FUNCTION_BLOCK SKILL_RunLogic (* The state machine of SKILL_Run: the precondition, waiting for the equipment, the command, the end condition, the timeout, the closing command. Technical: One run of a skill primitive: Pre, then the equipment free (0.5 s grace), Command until Post or the timer (Timed), Inv over it, StopCommand at the end, played before the end is reported *)
  (* Standard: 61499-2 *)
  (* Version 0.1, 2026-09-28, Project contributors, AAU Smart Production Lab *)
  PACKAGE modlib;
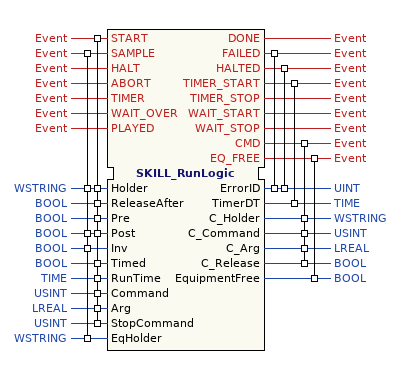
  EVENT_INPUT
    START WITH Holder, ReleaseAfter, Pre, Post, Timed, RunTime, Command, Arg, StopCommand; (* Start the run with what the contract says (Pre first) *)
    SAMPLE WITH Holder, Post, Inv, EqHolder; (* The equipment's newest state, as the contract judges it (Post, Inv, EqHolder) *)
    HALT; (* Stop the run (ErrorID Interrupted) *)
    ABORT; (* Abort the run: the equipment off and given up *)
    TIMER; (* The run's timer expired *)
    WAIT_OVER; (* Waited long enough for another holder to let go *)
    PLAYED; (* The command's phases were played *)
  END_EVENT
  EVENT_OUTPUT
    DONE; (* The run succeeded *)
    FAILED WITH ErrorID; (* The run failed (ErrorID) *)
    HALTED WITH ErrorID; (* The run was stopped *)
    TIMER_START WITH TimerDT; (* Start the timer (TimerDT) *)
    TIMER_STOP; (* Stop the timer *)
    WAIT_START; (* Start waiting for the equipment *)
    WAIT_STOP; (* Stop waiting *)
    CMD WITH C_Holder, C_Command, C_Arg, C_Release; (* Send a command to the equipment *)
    EQ_FREE WITH EquipmentFree; (* EquipmentFree is updated *)
  END_EVENT
  VAR_INPUT
    Holder : WSTRING; (* The name the equipment is held under: the skill's own, or for a step the skill it belongs to *)
    ReleaseAfter : BOOL; (* Give up the equipment with the run's last command *)
    Pre : BOOL; (* The precondition holds: the run may start (else PreconditionViolated, 1) *)
    Post : BOOL; (* The postcondition holds: the skill is done *)
    Inv : BOOL := TRUE; (* The invariant holds: the run may go on (else InvariantViolated, 2) *)
    Timed : BOOL; (* The skill ends after RunTime (TRUE), or when Post holds, failing after RunTime (FALSE) *)
    RunTime : TIME; (* How long it runs (Timed), or may take before it fails with Timeout (3) *)
    Command : USINT; (* The command's code to send while it runs *)
    Arg : LREAL; (* The command's argument (e.g. a position) *)
    StopCommand : USINT; (* The command's code to send when it is done or halted *)
    EqHolder : WSTRING; (* Who holds the equipment now (empty: free) *)
  END_VAR
  VAR_OUTPUT
    ErrorID : UINT; (* Error code: 0 none, 1 PreconditionViolated, 2 InvariantViolated, 3 Timeout, 4 NotReady, 5 NotPermitted, 6 Busy, 7 Interrupted, 8 OutOfRange *)
    TimerDT : TIME; (* How long the timer runs *)
    C_Holder : WSTRING; (* Sent with the command: who holds the equipment *)
    C_Command : USINT; (* Sent with the command: the command's code *)
    C_Arg : LREAL; (* Sent with the command: its argument (e.g. a position) *)
    C_Release : BOOL; (* Sent with the command: give up the equipment after it *)
    EquipmentFree : BOOL; (* The equipment is free, or held under Holder *)
  END_VAR
  VAR
    Outcome : USINT;
  END_VAR
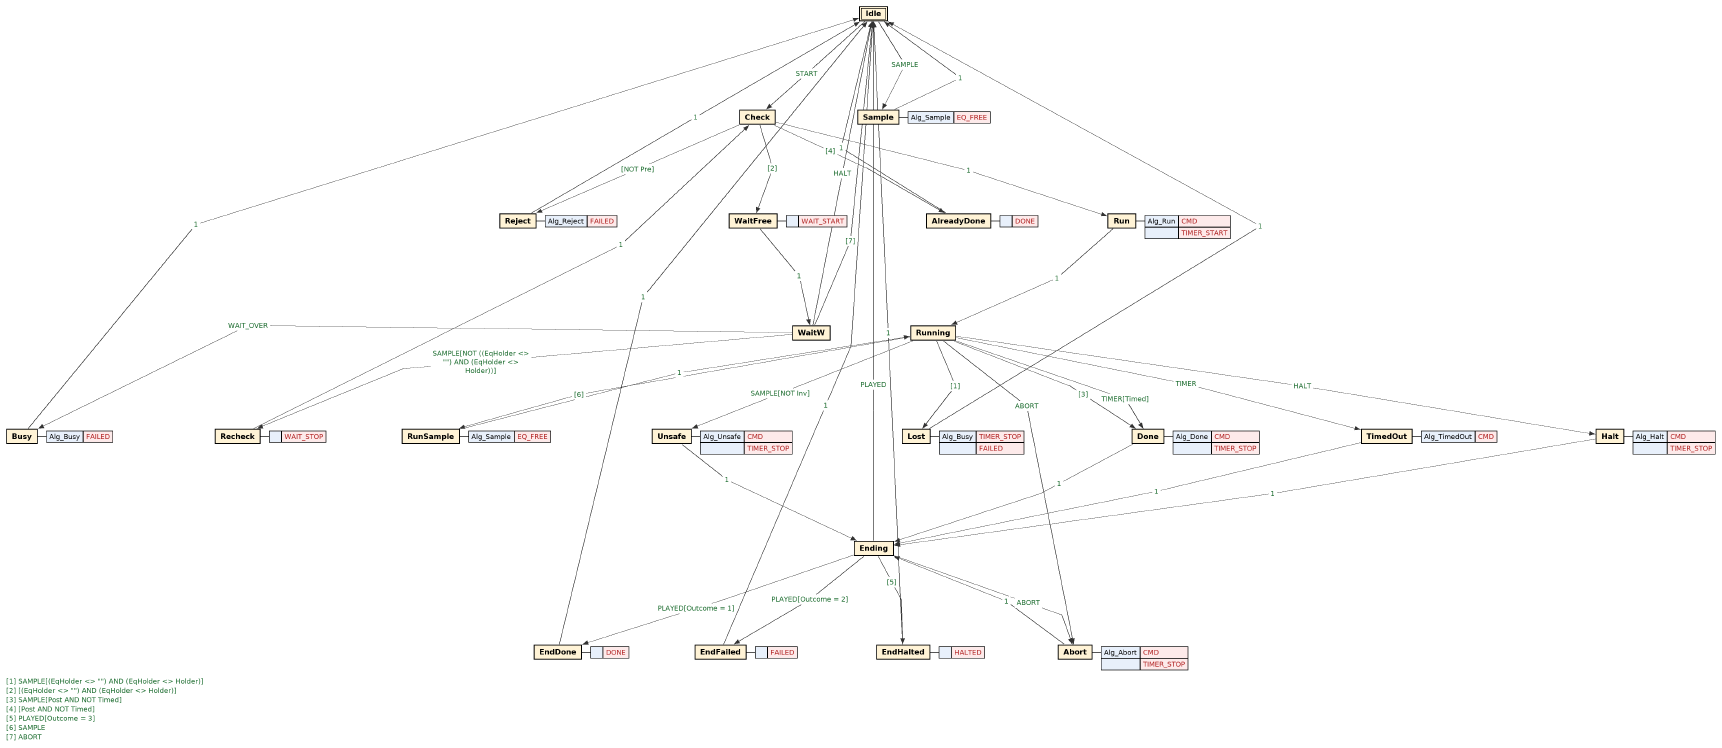
  EC_STATES
    Idle;
    Check;
    Reject : Alg_Reject -> FAILED;
    Sample : Alg_Sample -> EQ_FREE;
    Busy : Alg_Busy -> FAILED;
    WaitFree : -> WAIT_START;
    WaitW;
    Recheck : -> WAIT_STOP;
    AlreadyDone : -> DONE;
    Run : Alg_Run -> CMD, -> TIMER_START;
    RunSample : Alg_Sample -> EQ_FREE;
    Unsafe : Alg_Unsafe -> CMD, -> TIMER_STOP;
    Lost : Alg_Busy -> TIMER_STOP, -> FAILED;
    Done : Alg_Done -> CMD, -> TIMER_STOP;
    TimedOut : Alg_TimedOut -> CMD;
    Halt : Alg_Halt -> CMD, -> TIMER_STOP;
    Abort : Alg_Abort -> CMD, -> TIMER_STOP;
    Ending;
    EndDone : -> DONE;
    EndFailed : -> FAILED;
    EndHalted : -> HALTED;
    Running;
  END_STATES
  EC_TRANSITIONS
    Idle TO Check := START;
    Idle TO Sample := SAMPLE;
    Sample TO Idle := 1;
    Check TO Reject := [NOT Pre];
    Check TO WaitFree := [(EqHolder <> "") AND (EqHolder <> Holder)];
    WaitFree TO WaitW := 1;
    WaitW TO Recheck := SAMPLE[NOT ((EqHolder <> "") AND (EqHolder <> Holder))];
    WaitW TO Busy := WAIT_OVER;
    WaitW TO Idle := HALT;
    WaitW TO Idle := ABORT;
    Recheck TO Check := 1;
    Check TO AlreadyDone := [Post AND NOT Timed];
    Check TO Run := 1;
    Run TO Running := 1;
    Running TO Unsafe := SAMPLE[NOT Inv];
    Running TO Lost := SAMPLE[(EqHolder <> "") AND (EqHolder <> Holder)];
    Running TO Done := SAMPLE[Post AND NOT Timed];
    Running TO Done := TIMER[Timed];
    Running TO TimedOut := TIMER;
    Running TO RunSample := SAMPLE;
    RunSample TO Running := 1;
    Running TO Halt := HALT;
    Running TO Abort := ABORT;
    Reject TO Idle := 1;
    Busy TO Idle := 1;
    Lost TO Idle := 1;
    AlreadyDone TO Idle := 1;
    Unsafe TO Ending := 1;
    Done TO Ending := 1;
    TimedOut TO Ending := 1;
    Halt TO Ending := 1;
    Abort TO Ending := 1;
    Ending TO EndDone := PLAYED[Outcome = 1];
    Ending TO EndFailed := PLAYED[Outcome = 2];
    Ending TO EndHalted := PLAYED[Outcome = 3];
    Ending TO Idle := PLAYED;
    Ending TO Abort := ABORT;
    EndDone TO Idle := 1;
    EndFailed TO Idle := 1;
    EndHalted TO Idle := 1;
  END_TRANSITIONS
  ALGORITHM Alg_Reject IN ST:
ErrorID := 1;
  END_ALGORITHM
  ALGORITHM Alg_Sample IN ST:
EquipmentFree := (EqHolder = "") OR (EqHolder = Holder);
  END_ALGORITHM
  ALGORITHM Alg_Busy IN ST:
ErrorID := 6;
  END_ALGORITHM
  ALGORITHM Alg_Run IN ST:
C_Holder := Holder;
C_Command := Command;
C_Arg := Arg;
C_Release := FALSE;
TimerDT := RunTime;
  END_ALGORITHM
  ALGORITHM Alg_Unsafe IN ST:
C_Holder := Holder;
C_Command := 0;
C_Arg := Arg;
C_Release := ReleaseAfter;
ErrorID := 2;
Outcome := 2;
  END_ALGORITHM
  ALGORITHM Alg_Done IN ST:
C_Holder := Holder;
C_Command := StopCommand;
C_Arg := Arg;
C_Release := ReleaseAfter;
Outcome := 1;
  END_ALGORITHM
  ALGORITHM Alg_TimedOut IN ST:
C_Holder := Holder;
C_Command := 0;
C_Arg := Arg;
C_Release := ReleaseAfter;
ErrorID := 3;
Outcome := 2;
  END_ALGORITHM
  ALGORITHM Alg_Halt IN ST:
C_Holder := Holder;
C_Command := StopCommand;
C_Arg := Arg;
C_Release := ReleaseAfter;
ErrorID := 7;
Outcome := 3;
  END_ALGORITHM
  ALGORITHM Alg_Abort IN ST:
C_Holder := Holder;
C_Command := 0;
C_Arg := Arg;
C_Release := TRUE;
Outcome := 0;
  END_ALGORITHM
END_FUNCTION_BLOCK
